SUBAPPLICATION logiBUS_IXA_TO_PUBLISH_OPC (* Digitaler Eingang, lokaler OPC-UA-Write (ACTION=WRITE ohne Endpunkt) per AX_PUBLISH_1 *)
  (* Standard: 61499-2; Description: Copyright (c) 2026 Meisterschulen am Ostbahnhof This program and the accompanying materials are made available under the terms of the Eclipse Public License 2.0 which is available at https://www.eclipse.org/legal/epl-2.0/ SPDX-License-Identifier: EPL-2.0 *)
  (* Version 1.2, 2026-10-18, Franz Höpfinger, Meisterschulen am Ostbahnhof, Lokale Variante von logiBUS_IXA_TO_CLIENT_OPC: AX_PUBLISH_1 statt AX_CLIENT_1_0 *)
  (* Version 1.1, 2026-09-18, Franz Höpfinger, Meisterschulen am Ostbahnhof, logiBUS_IXA.INITO auf logiBUS_IXA.REQ zurueckverdrahtet (Selfloop) - loest nach der Initialisierung sofort einen Service-Request aus, statt auf die erste echte Wertaenderung am Bus zu warten (Fix fuer 'Waiting for handle'-Status direkt nach Boot). *)
  (* Version 1.0, 2026-09-02, Franz Höpfinger, Meisterschulen am Ostbahnhof, initial API and implementation and/or initial documentation *)
  PACKAGE MyLib::sys;
  IMPORT logiBUS::io::DI::logiBUS_DI;
  IMPORT logiBUS::io::DI::logiBUS_DI_S;
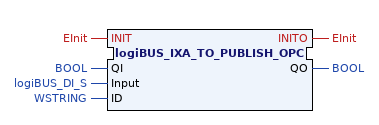
  EVENT_INPUT
    INIT : EInit; (* Initialization Request *)
  END_EVENT
  EVENT_OUTPUT
    INITO : EInit; (* Initialization Confirm *)
  END_EVENT
  VAR_INPUT
    QI : BOOL := TRUE; (* Quality Input - TRUE to enable service *)
    Input : logiBUS::io::DI::logiBUS_DI_S := logiBUS_DI::Invalid; (* Identify the Input Input_I1..I8 *)
    ID : WSTRING; (* Lokale Knotenadresse (BOOL, ACTION=WRITE, ohne Endpunkt) *)
  END_VAR
  VAR_OUTPUT
    QO : BOOL; (* Quality Output - TRUE if service executed successfully *)
  END_VAR
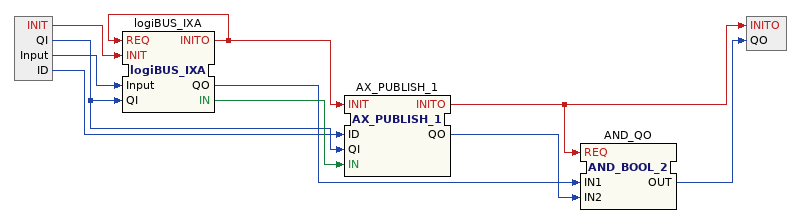
  FBS
    logiBUS_IXA : logiBUS::io::DI::logiBUS_IXA;
    AX_PUBLISH_1 : adapter::net::AX_PUBLISH_1;
    AND_QO : iec61131::booleanOperators::AND_BOOL_2;
  END_FBS
  EVENT_CONNECTIONS
    logiBUS_IXA.INITO TO logiBUS_IXA.REQ;
    INIT TO logiBUS_IXA.INIT;
    logiBUS_IXA.INITO TO AX_PUBLISH_1.INIT;
    AX_PUBLISH_1.INITO TO INITO;
    AX_PUBLISH_1.INITO TO AND_QO.REQ;
  END_CONNECTIONS
  DATA_CONNECTIONS
    Input TO logiBUS_IXA.Input;
    ID TO AX_PUBLISH_1.ID;
    QI TO logiBUS_IXA.QI;
    QI TO AX_PUBLISH_1.QI;
    logiBUS_IXA.QO TO AND_QO.IN1;
    AX_PUBLISH_1.QO TO AND_QO.IN2;
    AND_QO.OUT TO QO;
  END_CONNECTIONS
  ADAPTER_CONNECTIONS
    logiBUS_IXA.IN TO AX_PUBLISH_1.IN;
  END_CONNECTIONS
END_SUBAPPLICATION
